(* IEC 61131-3 sources: 2026_Projet_YGO_ExcavatriceDragage/CODE_BACKUP/CODE_20260904_AvantWeekendBackup_v0.6.34/C_DIAG_RESEAUX, 5 files *)

(* ---- E_Diag_State.st ---- *)
(* =======================================================================
   📊 E_Diag_State — Enumération des états du cycle de diagnostic réseau
   ───────────────────────────────────────────────────────────────
   🎯 Rôle : Phases d'état de surveillance diagnostic d'un bus ou équipement
   📄 Doc métier : DOC/AF/AF_Partie-12_Fonction_Diagnostic_v1.4.md
   ======================================================================= *)
TYPE E_Diag_State :
(
    DISABLED   := 0,  (* Désactivé (surveillance non active) *)
    READY      := 1,  (* Opérationnel réel, pas de défaut *)
    INIT       := 2,  (* Initialisation / Recherche de réseau *)
    MONITORING := 3,  (* Surveillance active (états transitoires) *)
    ERROR      := 4,  (* Anomalie de communication *)
    SIMULATED  := 5   (* Bypass simulation ou bypass réseau IHM — pas le bus réel *)
);
END_TYPE

(* ---- ST_Diag_Device.st ---- *)
(* =======================================================================
   📊 ST_Diag_Device — Structure diagnostic d'un esclave ou bus
   ───────────────────────────────────────────────────────────────
   🎯 Rôle : Structure de donnees d'état, diagnostic et alarme d'un equipement réseau
   📄 Doc métier : DOC/AF/AF_Partie-12_Fonction_Diagnostic_v1.4.md
   ======================================================================= *)
TYPE ST_Diag_Device :
STRUCT
    Online         : BOOL;        (* Esclave visible sur le bus *)
    Operational    : BOOL;        (* Esclave en mode OP (opérationnel) *)
    Error          : BOOL;        (* Signal de défaut actif pour cet esclave *)
    ErrorId        : WORD;        (* Code défaut détaillé *)
    State          : E_Diag_State; (* Phase courante du cycle de diagnostic *)
    StateAtError   : E_Diag_State; (* Instantané de la phase lors de l'anomalie *)
END_STRUCT
END_TYPE

(* ---- FB_Diag_CanOpen.st ---- *)
(* =======================================================================
   📊 FB_Diag_CanOpen — Diagnostic bus CANopen & Esclave Joystick
   ───────────────────────────────────────────────────────────────
   🎯 Rôle : Surveillance bus CANopen master et esclave Joystick (Online/Op)
   🔌 Architecture : Publication ST_Diag_Device & E_Diag_State
   📄 Doc métier : DOC/AF/AF_Partie-12_Fonction_Diagnostic_v1.4.md
   ======================================================================= *)
FUNCTION_BLOCK PUBLIC FB_Diag_CanOpen
VAR_INPUT
    // === COMMANDES & CONTROLE ===
    Enable                      : BOOL;         // --> [CMD] Active la surveillance CAN
    Reset                       : BOOL;         // --> [CMD] Front d'acquittement des defauts

    // === ETATS BRUTS MATERIEL ===
    CANbusStateRaw              : INT;          // --> [HW]  Valeur brute CANbus.GetBusState() (2 = ACTIVE)
    DeviceJoystickStateRaw      : DEVICE_STATE; // --> [HW]  Valeur brute JOY1.GetDeviceState()

    // === BYPASS & SIMULATION ===
    SimBypassActive             : BOOL;         // --> [TST] TRUE = simulation active pour ce device
    NetworkBypassActive         : BOOL;         // --> [TST] TRUE = bypass reseau global IHM
    CanBusBypassActive          : BOOL;         // --> [TST] TRUE = bypass specifique bus CANopen maître
    JoystickBypassActive        : BOOL;         // --> [TST] TRUE = bypass specifique esclave Joystick
END_VAR
VAR_OUTPUT
    // === ETAT DU BLOC ===
    Ready                       : BOOL;         // <-- [STAT] Logique de surveillance active

    // === DIAGNOSTICS STRUCTURES PAR EQUIPEMENT ===
    DeviceCanOpenMaster         : ST_Diag_Device; // <-- [DIAG] Diagnostics bus CANopen maître (Online, Op, Error, ErrorId, State)
    DeviceJoystick              : ST_Diag_Device; // <-- [DIAG] Diagnostics esclave Joystick (Online, Op, Error, ErrorId, State)
END_VAR
VAR
    // === SOUS-INSTANCES FB ===
    ResetEdge                   : R_TRIG;       // * [INST] Detecteur front de reset

    // === CALCULS ET ETATS INTERNES ===
    CANbusOnlineReal            : BOOL;         // . [LOC]  Bus reellement actif, hors tout bypass
    DeviceJoystickOnlineReal    : BOOL;         // . [LOC]  Joystick reellement RUNNING, hors tout bypass
    CANbusOnlineEff             : BOOL;         // . [LOC]  Online effectif bus CAN (reel OU bypass)
    DeviceJoystickOnlineEff     : BOOL;         // . [LOC]  Operational effectif joystick (reel OU bypass)
END_VAR

{region "§1 Gate"}
// 🛑 1. GATE : Désactivation logique si Enable = FALSE
IF NOT Enable THEN
    Ready := FALSE;
    DeviceJoystick.State := E_Diag_State.DISABLED;
    DeviceJoystick.Online := FALSE;
    DeviceJoystick.Operational := FALSE;
    DeviceJoystick.Error := FALSE;
    DeviceJoystick.ErrorId := 16#0000;
    DeviceCanOpenMaster.State := E_Diag_State.DISABLED;
    DeviceCanOpenMaster.Online := FALSE;
    DeviceCanOpenMaster.Operational := FALSE;
    DeviceCanOpenMaster.Error := FALSE;
    DeviceCanOpenMaster.ErrorId := 16#0000;
    RETURN;
END_IF;

Ready := TRUE;
{endregion}

{region "§2 Interprétation valeurs brutes"}
// 🧮 2. INTERPRÉTATION DES VALEURS BRUTES
CANbusOnlineReal         := (CANbusStateRaw = 2);
DeviceJoystickOnlineReal := (DeviceJoystickStateRaw = DEVICE_STATE.RUNNING);

CANbusOnlineEff          := CANbusOnlineReal OR SimBypassActive OR NetworkBypassActive OR CanBusBypassActive;
DeviceJoystickOnlineEff  := DeviceJoystickOnlineReal OR SimBypassActive OR NetworkBypassActive OR JoystickBypassActive;
{endregion}

{region "§3 Reset front"}
// 🔑 3. RESET FRONT — Efface les défauts si la cause a disparu
ResetEdge(CLK := Reset);
IF ResetEdge.Q THEN
    IF (CANbusOnlineEff AND DeviceJoystickOnlineEff) THEN
        DeviceJoystick.ErrorId := 16#0000;
        DeviceJoystick.StateAtError := E_Diag_State.DISABLED;
    END_IF;
END_IF;
{endregion}

{region "§4 Diagnostic joystick"}
// 🔍 4. DIAGNOSTIC JOYSTICK
// Bit 0 : Perte de communication CAN
IF NOT CANbusOnlineEff THEN
    DeviceJoystick.ErrorId := DeviceJoystick.ErrorId OR 16#0001;  (* Perte liaison CAN joystick *)
ELSE
    DeviceJoystick.Online := TRUE;
    DeviceJoystick.ErrorId := DeviceJoystick.ErrorId AND 16#FFFE; (* Effacement auto si la liaison revient *)
END_IF;

// Bit 1 : Mode non-opérationnel (esclave CANopen en pré-op ou défaut)
IF NOT DeviceJoystickOnlineEff THEN
    DeviceJoystick.ErrorId := DeviceJoystick.ErrorId OR 16#0002;  (* Joystick pas opérationnel *)
    DeviceJoystick.Operational := FALSE;
ELSE
    DeviceJoystick.Operational := TRUE;
    DeviceJoystick.ErrorId := DeviceJoystick.ErrorId AND 16#FFFD; (* Effacement auto dès que RUNNING *)
END_IF;
{endregion}

{region "§5 Machine etat joystick"}
// 🚦 5. MACHINE D'ÉTAT JOYSTICK
IF DeviceJoystick.ErrorId <> 0 THEN
    DeviceJoystick.State := E_Diag_State.ERROR;
ELSIF NOT (DeviceJoystick.Online AND DeviceJoystick.Operational) THEN
    DeviceJoystick.State := E_Diag_State.INIT;
ELSIF (SimBypassActive OR NetworkBypassActive OR JoystickBypassActive) AND NOT (CANbusOnlineReal AND DeviceJoystickOnlineReal) THEN
    DeviceJoystick.State := E_Diag_State.SIMULATED;
ELSE
    DeviceJoystick.State := E_Diag_State.READY;
END_IF;
{endregion}

{region "§6 Sorties globales"}
// 📤 6. SORTIES GLOBALES
DeviceJoystick.Error := (DeviceJoystick.ErrorId <> 0);

DeviceCanOpenMaster.Operational := CANbusOnlineEff;
DeviceCanOpenMaster.Online := CANbusOnlineEff;
DeviceCanOpenMaster.Error := NOT CANbusOnlineEff;

IF NOT CANbusOnlineEff THEN
    DeviceCanOpenMaster.ErrorId := 16#0001;
    DeviceCanOpenMaster.State := E_Diag_State.ERROR;
    IF DeviceCanOpenMaster.StateAtError = E_Diag_State.DISABLED THEN
        DeviceCanOpenMaster.StateAtError := E_Diag_State.INIT;
    END_IF;
ELSIF (SimBypassActive OR NetworkBypassActive OR CanBusBypassActive) AND NOT CANbusOnlineReal THEN
    DeviceCanOpenMaster.ErrorId := 16#0000;
    DeviceCanOpenMaster.State := E_Diag_State.SIMULATED;
ELSE
    DeviceCanOpenMaster.ErrorId := 16#0000;
    DeviceCanOpenMaster.State := E_Diag_State.READY;
END_IF;
{endregion}

(* ---- FB_Diag_Ethercat.st ---- *)
(* =======================================================================
   📊 FB_Diag_Ethercat — Diagnostic bus EtherCAT & Esclaves (M3, COD1, COD2)
   ───────────────────────────────────────────────────────────────
   🎯 Rôle : Surveillance bus EtherCAT master, variateur M3 et codeurs M1/M2
   🔌 Architecture : Publication ST_Diag_Device par esclave & E_Diag_State
   📄 Doc métier : DOC/AF/AF_Partie-12_Fonction_Diagnostic_v1.4.md
   ======================================================================= *)
FUNCTION_BLOCK PUBLIC FB_Diag_Ethercat
VAR_INPUT
    // === COMMANDES & CONTROLE ===
    Enable                      : BOOL;         // --> [CMD] Active la surveillance EtherCAT
    Reset                       : BOOL;         // --> [CMD] Front d'acquittement des defauts

    // === ETATS BRUTS MATERIEL & BYPASS VARIATEUR M3 ===
    DeviceVariateurStateRaw     : DEVICE_STATE; // --> [HW]  Valeur brute AC600_ECAT_Drive.GetDeviceState()
    DeviceVariateurSimBypass    : BOOL;         // --> [TST] TRUE = simulation active variateur M3

    // === ETATS BRUTS MATERIEL & BYPASS ENCODEUR M1 ===
    DeviceEncoderM1StateRaw     : DEVICE_STATE; // --> [HW]  Valeur brute COD1_CODEUR.GetDeviceState()
    DeviceEncoderM1SimBypass    : BOOL;         // --> [TST] TRUE = simulation active encodeur M1

    // === ETATS BRUTS MATERIEL & BYPASS ENCODEUR M2 ===
    DeviceEncoderM2StateRaw     : DEVICE_STATE; // --> [HW]  Valeur brute COD2_CODEUR.GetDeviceState()
    DeviceEncoderM2SimBypass    : BOOL;         // --> [TST] TRUE = simulation active encodeur M2

    // === BYPASS RESEAU IHM & GRANULAIRES ===
    NetworkBypassActive         : BOOL;         // --> [TST] TRUE = bypass reseau global IHM
    EcatBusBypassActive         : BOOL;         // --> [TST] TRUE = bypass specifique bus EtherCAT maître
    VariateurBypassActive       : BOOL;         // --> [TST] TRUE = bypass specifique esclave variateur M3
    EncoderM1BypassActive       : BOOL;         // --> [TST] TRUE = bypass specifique esclave codeur M1
    EncoderM2BypassActive       : BOOL;         // --> [TST] TRUE = bypass specifique esclave codeur M2
END_VAR
VAR_OUTPUT
    // === ETAT DU BLOC ===
    Ready                       : BOOL;         // <-- [STAT] Logique de surveillance active

    // === DIAGNOSTICS STRUCTURES PAR EQUIPEMENT ===
    DeviceEthercatMaster        : ST_Diag_Device; // <-- [DIAG] Diagnostics bus EtherCAT
    DeviceVariateur             : ST_Diag_Device; // <-- [DIAG] Diagnostics esclave AC600
    DeviceEncoderM1             : ST_Diag_Device; // <-- [DIAG] Diagnostics esclave COD1
    DeviceEncoderM2             : ST_Diag_Device; // <-- [DIAG] Diagnostics esclave COD2
END_VAR
VAR
    // === SOUS-INSTANCES FB ===
    ResetEdge                   : R_TRIG;       // * [INST] Detecteur front de reset

    // === CALCULS ET ETATS INTERNES ===
    VariateurOnlineReal         : BOOL;         // . [LOC]  GetDeviceState() = RUNNING, hors tout bypass
    EncoderM1OnlineReal         : BOOL;         // . [LOC]  GetDeviceState() = RUNNING, hors tout bypass
    EncoderM2OnlineReal         : BOOL;         // . [LOC]  GetDeviceState() = RUNNING, hors tout bypass
    VariateurBypass             : BOOL;         // . [LOC]  Simulation OU bypass reseau IHM variateur
    EncoderM1Bypass             : BOOL;         // . [LOC]  Simulation OU bypass reseau IHM encodeur M1
    EncoderM2Bypass             : BOOL;         // . [LOC]  Simulation OU bypass reseau IHM encodeur M2
    VariateurOnlineEff          : BOOL;         // . [LOC]  Online effectif (reel OU bypass)
    EncoderM1OnlineEff          : BOOL;         // . [LOC]  Online effectif (reel OU bypass)
    EncoderM2OnlineEff          : BOOL;         // . [LOC]  Online effectif (reel OU bypass)
END_VAR

{region "§1 Gate de desactivation"}
// 🛑 1. GATE : Désactivation si Enable = FALSE
IF NOT Enable THEN
    Ready := FALSE;
    DeviceVariateur.State := E_Diag_State.DISABLED;
    DeviceEncoderM1.State := E_Diag_State.DISABLED;
    DeviceEncoderM2.State := E_Diag_State.DISABLED;
    DeviceVariateur.Online := FALSE;
    DeviceEncoderM1.Online := FALSE;
    DeviceEncoderM2.Online := FALSE;
    DeviceVariateur.Operational := FALSE;
    DeviceEncoderM1.Operational := FALSE;
    DeviceEncoderM2.Operational := FALSE;
    DeviceVariateur.Error := FALSE;
    DeviceEncoderM1.Error := FALSE;
    DeviceEncoderM2.Error := FALSE;
    DeviceEthercatMaster.State := E_Diag_State.DISABLED;
    DeviceEthercatMaster.Online := FALSE;
    DeviceEthercatMaster.Operational := FALSE;
    DeviceEthercatMaster.Error := FALSE;
    DeviceEthercatMaster.ErrorId := 16#0000;
    RETURN;
END_IF;

Ready := TRUE;

{endregion}

{region "§2 Interpretation etats bruts et bypass"}
// 🧮 2. INTERPRÉTATION DES VALEURS BRUTES
VariateurOnlineReal := (DeviceVariateurStateRaw = DEVICE_STATE.RUNNING);
EncoderM1OnlineReal := (DeviceEncoderM1StateRaw = DEVICE_STATE.RUNNING);
EncoderM2OnlineReal := (DeviceEncoderM2StateRaw = DEVICE_STATE.RUNNING);

VariateurBypass := DeviceVariateurSimBypass OR NetworkBypassActive OR VariateurBypassActive;
EncoderM1Bypass := DeviceEncoderM1SimBypass OR NetworkBypassActive OR EncoderM1BypassActive;
EncoderM2Bypass := DeviceEncoderM2SimBypass OR NetworkBypassActive OR EncoderM2BypassActive;

VariateurOnlineEff := VariateurOnlineReal OR VariateurBypass;
EncoderM1OnlineEff := EncoderM1OnlineReal OR EncoderM1Bypass;
EncoderM2OnlineEff := EncoderM2OnlineReal OR EncoderM2Bypass;

// 🔑 3. RESET FRONT
ResetEdge(CLK := Reset);

{endregion}

{region "§3 Diagnostic par equipement"}
// 🔍 4. DIAGNOSTIC VARIATEUR (AC600_ECAT_Drive / Translation M3)
DeviceVariateur.Online := VariateurOnlineEff;
DeviceVariateur.Operational := VariateurOnlineEff;

IF NOT DeviceVariateur.Online THEN
    DeviceVariateur.ErrorId := DeviceVariateur.ErrorId OR 16#0010;  (* Perte liaison physique variateur *)
ELSE
    DeviceVariateur.ErrorId := DeviceVariateur.ErrorId AND 16#FFEF; (* Effacement auto dès que RUNNING *)
END_IF;

// 🔍 5. DIAGNOSTIC ENCODEUR M1 (COD1_CODEUR / WinchM1)
DeviceEncoderM1.Online := EncoderM1OnlineEff;
DeviceEncoderM1.Operational := EncoderM1OnlineEff;

IF NOT DeviceEncoderM1.Online THEN
    DeviceEncoderM1.ErrorId := DeviceEncoderM1.ErrorId OR 16#0020;  (* Perte liaison encodeur M1 *)
ELSE
    DeviceEncoderM1.ErrorId := DeviceEncoderM1.ErrorId AND 16#FFDF; (* Effacement auto dès que RUNNING *)
END_IF;

// 🔍 6. DIAGNOSTIC ENCODEUR M2 (COD2_CODEUR / WinchM2)
DeviceEncoderM2.Online := EncoderM2OnlineEff;
DeviceEncoderM2.Operational := EncoderM2OnlineEff;

IF NOT DeviceEncoderM2.Online THEN
    DeviceEncoderM2.ErrorId := DeviceEncoderM2.ErrorId OR 16#0030;  (* Perte liaison encodeur M2 *)
ELSE
    DeviceEncoderM2.ErrorId := DeviceEncoderM2.ErrorId AND 16#FFCF; (* Effacement auto dès que RUNNING *)
END_IF;

{endregion}

{region "§4 Etats diagnostic par equipement"}
// 🚦 7. STATE MACHINES DE CHAQUE APPAREIL
IF DeviceVariateur.ErrorId <> 0 THEN
    DeviceVariateur.State := E_Diag_State.ERROR;
ELSIF NOT VariateurOnlineEff THEN
    DeviceVariateur.State := E_Diag_State.INIT;
ELSIF VariateurBypass AND NOT VariateurOnlineReal THEN
    DeviceVariateur.State := E_Diag_State.SIMULATED;
ELSE
    DeviceVariateur.State := E_Diag_State.READY;
END_IF;

IF DeviceEncoderM1.ErrorId <> 0 THEN
    DeviceEncoderM1.State := E_Diag_State.ERROR;
ELSIF NOT EncoderM1OnlineEff THEN
    DeviceEncoderM1.State := E_Diag_State.INIT;
ELSIF EncoderM1Bypass AND NOT EncoderM1OnlineReal THEN
    DeviceEncoderM1.State := E_Diag_State.SIMULATED;
ELSE
    DeviceEncoderM1.State := E_Diag_State.READY;
END_IF;

IF DeviceEncoderM2.ErrorId <> 0 THEN
    DeviceEncoderM2.State := E_Diag_State.ERROR;
ELSIF NOT EncoderM2OnlineEff THEN
    DeviceEncoderM2.State := E_Diag_State.INIT;
ELSIF EncoderM2Bypass AND NOT EncoderM2OnlineReal THEN
    DeviceEncoderM2.State := E_Diag_State.SIMULATED;
ELSE
    DeviceEncoderM2.State := E_Diag_State.READY;
END_IF;

{endregion}

{region "§5 Synthese EtherCAT et sorties"}
// 📤 8. RÉSUMÉ ET DÉFAUTS
DeviceVariateur.Error := (DeviceVariateur.ErrorId <> 0);
DeviceEncoderM1.Error := (DeviceEncoderM1.ErrorId <> 0);
DeviceEncoderM2.Error := (DeviceEncoderM2.ErrorId <> 0);

DeviceEthercatMaster.Online := (VariateurOnlineEff AND EncoderM1OnlineEff AND EncoderM2OnlineEff) OR NetworkBypassActive OR EcatBusBypassActive;
DeviceEthercatMaster.Operational := DeviceEthercatMaster.Online;
DeviceEthercatMaster.Error := NOT DeviceEthercatMaster.Operational;

IF DeviceEthercatMaster.Error THEN
    DeviceEthercatMaster.ErrorId := 16#0001;
    DeviceEthercatMaster.State := E_Diag_State.ERROR;
ELSIF (VariateurBypass OR EncoderM1Bypass OR EncoderM2Bypass OR EcatBusBypassActive) THEN
    DeviceEthercatMaster.ErrorId := 16#0000;
    DeviceEthercatMaster.State := E_Diag_State.SIMULATED;
ELSE
    DeviceEthercatMaster.ErrorId := 16#0000;
    DeviceEthercatMaster.State := E_Diag_State.READY;
END_IF;
{endregion}

(* ---- FB_Diag_IhmHeartbeat.st ---- *)
(* =======================================================================
   📊 FB_Diag_IhmHeartbeat — Surveillance bidirectionnelle Heartbeat IHM/PLC
   ───────────────────────────────────────────────────────────────
   🎯 Rôle : Surveillance toggle IHM, generation toggle PLC et diagnostic timeout
   🛡️ Protection : FB de diagnostic autonome (sans action directe sur AU)
   📄 Doc métier : DOC/AF/AF_Partie-12_Fonction_Diagnostic_v1.4.md
   ======================================================================= *)
FUNCTION_BLOCK PUBLIC FB_Diag_IhmHeartbeat
VAR_INPUT
    // === COMMANDES & REGLAGES ===
    Enable                      : BOOL;         // --> [CMD] Active la surveillance (FALSE = IHM invalide)
    TglHeartbeatIhm             : BOOL;         // --> [HW]  Toggle IHM, inversion attendue toutes les 500 ms
    IhmTimeout                  : TIME := T#2s; // --> [CFG] Absence maximale de front IHM
    PlcTogglePeriod             : TIME := T#500ms; // --> [CFG] Periode du clignotant PLC
END_VAR
VAR_OUTPUT
    // === ETATS & DIAGNOSTICS IHM ===
    HeartbeatIhmOk              : BOOL;         // <-- [STAT] TRUE apres front IHM post-boot et avant timeout
    HeartbeatIhmTimeout         : BOOL;         // <-- [DIAG] TRUE = aucun front IHM depuis IhmTimeout
    TglHeartbeatPlc             : BOOL;         // <-- [STAT] Clignotant PLC a superviser cote IHM
    TimeSinceIhmEdge            : TIME;         // <-- [DIAG] Temps ecoule depuis le dernier front IHM
END_VAR
VAR
    // === SOUS-INSTANCES FB ===
    IhmTimeoutTon               : TON;          // * [INST] Timer de surveillance timeout IHM
    PlcToggleTon                : TON;          // * [INST] Timer clignotant heartbeat PLC

    // === CALCULS ET ETATS INTERNES ===
    LastIhmToggle               : BOOL;         // . [LOC]  Memoire du dernier etat toggle IHM
    IhmEdgeSeen                 : BOOL;         // . [LOC]  Verrou front vu (interdit RETAIN au boot)
    IhmEdgeDetected             : BOOL;         // . [LOC]  Front de changement toggle IHM detecte
END_VAR

// === IMPLEMENTATION ===

{region "§1 Gate"}
// 🛑 Sans Enable, aucune valeur mémorisée ne peut déclarer l'IHM valide.
IF NOT Enable THEN
    HeartbeatIhmOk := FALSE;
    HeartbeatIhmTimeout := TRUE;
    TglHeartbeatPlc := FALSE;
    TimeSinceIhmEdge := T#0s;
    LastIhmToggle := TglHeartbeatIhm;
    IhmEdgeSeen := FALSE;
    IhmTimeoutTon(IN := FALSE, PT := IhmTimeout);
    PlcToggleTon(IN := FALSE, PT := PlcTogglePeriod);
    RETURN;
END_IF;
{endregion}

{region "§2 Front IHM"}
// 📥 Front par comparaison : l'IHM écrit un BOOL toggle, pas une impulsion courte.
IhmEdgeDetected := (TglHeartbeatIhm <> LastIhmToggle);
LastIhmToggle := TglHeartbeatIhm;
IF IhmEdgeDetected THEN
    IhmEdgeSeen := TRUE;
END_IF;
{endregion}

{region "§3 Timeout IHM"}
// ⏱️ Le timer repart à chaque front. Au boot, il atteint le timeout au bout de IhmTimeout.
// HeartbeatIhmOk reste TRUE tant que le timeout n'est pas expiré (boot propre sans alarme au scan 1).
IhmTimeoutTon(IN := NOT IhmEdgeDetected, PT := IhmTimeout);
TimeSinceIhmEdge := IhmTimeoutTon.ET;
HeartbeatIhmTimeout := IhmTimeoutTon.Q;
HeartbeatIhmOk := NOT HeartbeatIhmTimeout;
{endregion}

{region "§4 Clignotant PLC"}
// 💡 Clignotant PLC indépendant : information de vie pour l'IHM, jamais signal Signal Safety autonome.
PlcToggleTon(IN := NOT PlcToggleTon.Q, PT := PlcTogglePeriod);
IF PlcToggleTon.Q THEN
    TglHeartbeatPlc := NOT TglHeartbeatPlc;
END_IF;
{endregion}
